TYPE "DT_MEASUREMENT_SYSTEM_GENERATOR_EXCITATION"
VERSION : 0.1
   STRUCT
      I_1 { S7_SetPoint := 'False'} : "DT_MEASUREMENT_SOLO" := ((), (), FALSE, 1, 0, 96, 32000, 32000, 32000, 0, 0, 0, 0, 0, 0, 0, 0, 0, 0, 0, 0, 0, 0.0, '');
      I_2 { S7_SetPoint := 'False'} : "DT_MEASUREMENT_SOLO" := ((), (), FALSE, 1, 0, 97, 32000, 32000, 32000, 0, 0, 0, 0, 0, 0, 0, 0, 0, 0, 0, 0, 0, 0.0, '');
      I_3 { S7_SetPoint := 'False'} : "DT_MEASUREMENT_SOLO" := ((), (), FALSE, 1, 0, 98, 32000, 32000, 32000, 0, 0, 0, 0, 0, 0, 0, 0, 0, 0, 0, 0, 0, 0.0, '');
      I { S7_SetPoint := 'False'} : "DT_MEASUREMENT_SOLO" := ((), (), FALSE, 1, 0, 99, 32000, 32000, 32000, 0, 0, 0, 0, 0, 0, 0, 0, 0, 0, 0, 0, 0, 0.0, '');
      U12 { S7_SetPoint := 'False'} : "DT_MEASUREMENT_SOLO" := ((), (), FALSE, 1, 0, 100, 32000, 32000, 32000, 0, 0, 0, 0, 0, 0, 0, 0, 0, 0, 0, 0, 0, 0.0, '');
      U13 { S7_SetPoint := 'False'} : "DT_MEASUREMENT_SOLO" := ((), (), FALSE, 1, 0, 101, 32000, 32000, 32000, 0, 0, 0, 0, 0, 0, 0, 0, 0, 0, 0, 0, 0, 0.0, '');
      U23 { S7_SetPoint := 'False'} : "DT_MEASUREMENT_SOLO" := ((), (), FALSE, 1, 0, 102, 32000, 32000, 32000, 0, 0, 0, 0, 0, 0, 0, 0, 0, 0, 0, 0, 0, 0.0, '');
      U_LL { S7_SetPoint := 'False'} : "DT_MEASUREMENT_SOLO" := ((), (), FALSE, 1, 0, 103, 32000, 32000, 32000, 0, 0, 0, 0, 0, 0, 0, 0, 0, 0, 0, 0, 0, 0.0, '');
      Field_current { S7_SetPoint := 'False'} : "DT_MEASUREMENT_SOLO" := ((), (), FALSE, 1, 0, 104, 32000, 32000, 32000, 0, 0, 0, 0, 0, 0, 0, 0, 0, 0, 0, 0, 0, 0.0, '');
      Field_voltage { S7_SetPoint := 'False'} : "DT_MEASUREMENT_SOLO" := ((), (), FALSE, 1, 0, 105, 32000, 32000, 32000, 0, 0, 0, 0, 0, 0, 0, 0, 0, 0, 0, 0, 0, 0.0, '');
      Auxiliary_current { S7_SetPoint := 'False'} : "DT_MEASUREMENT_SOLO" := ((), (), FALSE, 1, 0, 106, 32000, 32000, 32000, 0, 0, 0, 0, 0, 0, 0, 0, 0, 0, 0, 0, 0, 0.0, '');
      f { S7_SetPoint := 'False'} : "DT_MEASUREMENT_SOLO" := ((), (), FALSE, 1, 0, 107, 32000, 32000, 32000, 0, 0, 0, 0, 0, 0, 0, 0, 0, 0, 0, 0, 0, 0.0, '');
      PF { S7_SetPoint := 'False'} : "DT_MEASUREMENT_SOLO" := ((), (), FALSE, 1, 0, 108, 32000, 32000, 32000, 0, 0, 0, 0, 0, 0, 0, 0, 0, 0, 0, 0, 0, 0.0, '');
      P { S7_SetPoint := 'False'} : "DT_MEASUREMENT_SOLO" := ((), (), FALSE, 1, 0, 109, 32000, 32000, 32000, 0, 0, 0, 0, 0, 0, 0, 0, 0, 0, 0, 0, 0, 0.0, '');
      Q { S7_SetPoint := 'False'} : "DT_MEASUREMENT_SOLO" := ((), (), FALSE, 1, 0, 110, 32000, 32000, 32000, 0, 0, 0, 0, 0, 0, 0, 0, 0, 0, 0, 0, 0, 0.0, '');
      S { S7_SetPoint := 'False'} : "DT_MEASUREMENT_SOLO" := ((), (), FALSE, 1, 0, 111, 32000, 32000, 32000, 0, 0, 0, 0, 0, 0, 0, 0, 0, 0, 0, 0, 0, 0.0, '');
      E_ACT_IMP { S7_SetPoint := 'False'} : "DT_MEASUREMENT_SOLO" := ((), (), FALSE, 1, 0, 112, 32000, 32000, 32000, 0, 0, 0, 0, 0, 0, 0, 0, 0, 0, 0, 0, 0, 0.0, '');
      E_ACT_EXP { S7_SetPoint := 'False'} : "DT_MEASUREMENT_SOLO" := ((), (), FALSE, 1, 0, 113, 32000, 32000, 32000, 0, 0, 0, 0, 0, 0, 0, 0, 0, 0, 0, 0, 0, 0.0, '');
      E_RACT_IMP { S7_SetPoint := 'False'} : "DT_MEASUREMENT_SOLO" := ((), (), FALSE, 1, 0, 114, 32000, 32000, 32000, 0, 0, 0, 0, 0, 0, 0, 0, 0, 0, 0, 0, 0, 0.0, '');
      E_RACT_EXP { S7_SetPoint := 'False'} : "DT_MEASUREMENT_SOLO" := ((), (), FALSE, 1, 0, 115, 32000, 32000, 32000, 0, 0, 0, 0, 0, 0, 0, 0, 0, 0, 0, 0, 0, 0.0, '');
      Spare_1 { S7_SetPoint := 'False'} : "DT_MEASUREMENT_SOLO" := ((), (), FALSE, 1, 0, 116, 32000, 32000, 32000, 0, 0, 0, 0, 0, 0, 0, 0, 0, 0, 0, 0, 0, 0.0, '');
      Spare_2 { S7_SetPoint := 'False'} : "DT_MEASUREMENT_SOLO" := ((), (), FALSE, 1, 0, 117, 32000, 32000, 32000, 0, 0, 0, 0, 0, 0, 0, 0, 0, 0, 0, 0, 0, 0.0, '');
      Spare_3 { S7_SetPoint := 'False'} : "DT_MEASUREMENT_SOLO" := ((), (), FALSE, 1, 0, 118, 32000, 32000, 32000, 0, 0, 0, 0, 0, 0, 0, 0, 0, 0, 0, 0, 0, 0.0, '');
      Spare { S7_SetPoint := 'False'} : "DT_MEASUREMENT_SOLO" := ((), (), FALSE, 1, 0, 119, 32000, 32000, 32000, 0, 0, 0, 0, 0, 0, 0, 0, 0, 0, 0, 0, 0, 0.0, '');
   END_STRUCT;

END_TYPE

